(* IEC 61131-3 sources: iolistgen/tests_support/pl_stub/src/Interfaces/I_AlarmSink, 1 file *)

(* ---- OnAlarmEvent.method.decl.st ---- *)
METHOD OnAlarmEvent : BOOL
VAR_IN_OUT CONSTANT
    // lint:allow STL007 VAR_IN_OUT CONSTANT — ссылка только для чтения, а не константа (API.md, раздел 0)
    stEvent : ST_AlarmEvent;
END_VAR
